(* IEC 61131-3 sources: scada/02_Delta_PLC_HMI_ONTAS/kod, 2 files *)

(* ---- FB_AnalogOlcek.st ---- *)
(* ==========================================================================
   FB_AnalogOlcek - Analog giriş ölçekleme + filtre + kopuk kablo tespiti
   Delta AS/DVP analog modülü: 4-20 mA -> ham 0..32000 (modüle göre ayarlanır)
   ========================================================================== *)
FUNCTION_BLOCK FB_AnalogOlcek
VAR_INPUT
    HamDeger   : INT;            (* Modülden okunan ham değer *)
    HamMin     : INT  := 0;      (* 4 mA karşılığı *)
    HamMax     : INT  := 32000;  (* 20 mA karşılığı *)
    MuhMin     : REAL := 0.0;    (* Örn. 0 bar *)
    MuhMax     : REAL := 10.0;   (* Örn. 10 bar *)
    KopukLimit : INT  := -500;   (* 4 mA altı: kablo kopuk *)
END_VAR
VAR_OUTPUT
    Deger      : REAL;           (* Filtrelenmiş mühendislik değeri *)
    KopukAlarm : BOOL;
END_VAR
VAR
    Tampon     : ARRAY[0..9] OF REAL;
    Indeks     : INT;
    Toplam     : REAL;
    i          : INT;
    Anlik      : REAL;
END_VAR

KopukAlarm := HamDeger < KopukLimit;

(* Doğrusal ölçekleme: y = (x - x1) * (y2 - y1) / (x2 - x1) + y1 *)
Anlik := INT_TO_REAL(HamDeger - HamMin) * (MuhMax - MuhMin)
         / INT_TO_REAL(HamMax - HamMin) + MuhMin;

(* Sınırla *)
IF Anlik < MuhMin THEN Anlik := MuhMin; END_IF;
IF Anlik > MuhMax THEN Anlik := MuhMax; END_IF;

(* 10 örnekli hareketli ortalama *)
Tampon[Indeks] := Anlik;
Indeks := (Indeks + 1) MOD 10;
Toplam := 0.0;
FOR i := 0 TO 9 DO
    Toplam := Toplam + Tampon[i];
END_FOR;
Deger := Toplam / 10.0;

END_FUNCTION_BLOCK

(* ---- FB_MakineSekans.st ---- *)
(* ==========================================================================
   FB_MakineSekans - Adım (step) tabanlı otomatik makine çevrimi
   Besleme -> Sıkma -> İşlem -> Açma -> Boşaltma -> Başa dön
   ========================================================================== *)
FUNCTION_BLOCK FB_MakineSekans
VAR_INPUT
    Start, Stop, Reset   : BOOL;
    UrunVar              : BOOL;   (* Besleme sensörü *)
    SikmaIleri, SikmaGeri: BOOL;   (* Silindir manyetik sensörleri *)
    IslemSuresi          : TIME := T#3s;
    AdimZamanAsimi       : TIME := T#10s;
END_VAR
VAR_OUTPUT
    Y_Besleme, Y_Sikma, M_Islem, Y_Bosalt : BOOL;
    Adim     : INT;     (* HMI'da gösterilir *)
    Alarm    : BOOL;
    Sayac    : DINT;    (* Üretim sayacı *)
END_VAR
VAR
    Calisiyor : BOOL;
    tIslem    : TON;
    tAsim     : TON;
    OncekiAdim: INT;
END_VAR

IF Reset THEN Alarm := FALSE; Adim := 0; END_IF;
IF Stop OR Alarm THEN Calisiyor := FALSE; END_IF;
IF Start AND NOT Alarm THEN Calisiyor := TRUE; END_IF;

(* Her adımın zaman aşımı denetimi: adım değişince sayaç sıfırlanır *)
tAsim(IN := Calisiyor AND (Adim = OncekiAdim) AND (Adim <> 0), PT := AdimZamanAsimi);
OncekiAdim := Adim;
IF tAsim.Q THEN Alarm := TRUE; END_IF;

IF Calisiyor THEN
    CASE Adim OF
    0:  IF NOT UrunVar THEN Adim := 10; END_IF;           (* Yuva boş mu? *)
    10: Y_Besleme := TRUE;                                 (* Ürünü besle *)
        IF UrunVar THEN Y_Besleme := FALSE; Adim := 20; END_IF;
    20: Y_Sikma := TRUE;                                   (* Sık *)
        IF SikmaIleri THEN Adim := 30; END_IF;
    30: M_Islem := TRUE;                                   (* İşlem *)
        tIslem(IN := TRUE, PT := IslemSuresi);
        IF tIslem.Q THEN
            M_Islem := FALSE; tIslem(IN := FALSE); Adim := 40;
        END_IF;
    40: Y_Sikma := FALSE;                                  (* Aç *)
        IF SikmaGeri THEN Adim := 50; END_IF;
    50: Y_Bosalt := TRUE;                                  (* Boşalt *)
        IF NOT UrunVar THEN
            Y_Bosalt := FALSE; Sayac := Sayac + 1; Adim := 0;
        END_IF;
    END_CASE;
ELSE
    Y_Besleme := FALSE; M_Islem := FALSE; Y_Bosalt := FALSE;
END_IF;

END_FUNCTION_BLOCK
